// TIA Portal V21 export
DATA_BLOCK "IDB_AnaStatusIgnored"   // DB16
// stored: InstanceOfName FB_AnaStatusIgnored, InstanceOfType FB
"FB_AnaStatusIgnored"
   // VAR
   //    Now : DTL;
   // END_VAR
BEGIN
END_DATA_BLOCK
